(* IEC 61131-3 sources: Lasal-MCP/examples/SampleSource/2_PumpControlSolution/Stations/MachineControl/MachineControl/Class/SafetyBaseFSoE (part 3) *)

                b_NeedApplicationRestart := TRUE;
              end_if;
            end_if;
          end_if;
        end_if;

//*****************************************************************************
//**   UNSAFE BOOL INPUT VARIABLES                                           **
//*****************************************************************************

        // here we go for unsafe bool input vars

        // get number of unsafe input vars
        sd_retval := SDOReadCfgRequ ( p_SDORequestBuffer  := p_SDORequestBuffer
                                    , p_SDOResponseBuffer := p_SDOResponseBuffer
                                    , ud_Address          := ud_Address
                                    , us_Length           := 4
                                    );

        //no response
        if ( sd_retval <> 0 ) then
          LogError("@0217 (SafetyBaseFSoE::ReadSDOConfig) Config Read Error: Failed to read number of unsafe input vars.");
          return;
        end_if;

        ud_CntUnsafeInputs := p_SDOResponseBuffer^.ud_Data;

        ud_Address := p_SDORequestBuffer^.ud_Address + 4;

        // skip the names of unsafe inputs
        for i := 1 to ud_CntUnsafeInputs do

          // get length of Name
          sd_retval := SDOReadCfgRequ ( p_SDORequestBuffer  := p_SDORequestBuffer
                                      , p_SDOResponseBuffer := p_SDOResponseBuffer
                                      , ud_Address          := ud_Address
                                      , us_Length           := 4
                                      );
          //no response
          if ( sd_retval <> 0 ) then
            LogError("@0218 (SafetyBaseFSoE::ReadSDOConfig) Config Read Error: Reading length of unsafe input name failed.");
            return;
          end_if;

          // prepare address to get name
          ud_Address += 4;

//          ud_ActStrLen := ud_TmpStrLen := p_SDOResponseBuffer^.ud_Data;
          ud_TmpStrLen := p_SDOResponseBuffer^.ud_Data;
          ud_ActStrLen := ud_TmpStrLen;
          ud_TmpAddress := ud_Address;

          IF p_BlockedTransferMemory = NIL THEN
            sd_retval := -100;
            SetSafetyState(NewState:=_MemAllocFailed);
            RETURN;
          END_IF;

          IF ud_BlockedTransferMemorySize < (ud_TmpStrLen + 1) THEN
            p_BlockedTransferMemory := ToStdLib.ReAlloc(mptr:=p_BlockedTransferMemory, newsize:=GetNewMemSize(ud_TmpStrLen + 1));
            IF p_BlockedTransferMemory = NIL THEN
              ud_BlockedTransferMemorySize := 0;
              sd_retval := -100;
              SetSafetyState(NewState:=_MemAllocFailed);
              RETURN;
            ELSE
              ud_BlockedTransferMemorySize := GetNewMemSize(ud_TmpStrLen + 1);
            END_IF;
          END_IF;

          ToStdLib.MemSet(dest:=p_BlockedTransferMemory, value:=0, size:=ud_BlockedTransferMemorySize);

          p_TmpBlockedData := p_BlockedTransferMemory;

          us_BlockedTransferLength := BlockedTransferLength(ud_Datalength:=ud_TmpStrLen, us_MaxBlocklength:=60);

          while us_BlockedTransferLength do

            // get name
            sd_retval := SDOReadCfgRequ ( p_SDORequestBuffer  := p_SDORequestBuffer
                                        , p_SDOResponseBuffer := p_SDOResponseBuffer
                                        , ud_Address          := ud_TmpAddress
                                        , us_Length           := us_BlockedTransferLength
                                        , b_UseCache          := us_BlockedTransferLength < us_DataLength_Max
                                        );
            //no response
            if ( sd_retval <> 0 ) then
              LogError("@0219 (SafetyBaseFSoE::ReadSDOConfig) Config Read Error: Reading unsafe input name failed.");
              return;
            end_if;

            ToStdLib.MemCpy(dest:=p_TmpBlockedData,
                             source:=#p_SDOResponseBuffer^.ud_Data,
                             size:=us_BlockedTransferLength);

            p_TmpBlockedData += us_BlockedTransferLength;
            ud_TmpAddress += us_BlockedTransferLength;
            ud_TmpStrLen -= us_BlockedTransferLength;

            us_BlockedTransferLength := BlockedTransferLength(ud_Datalength:=ud_TmpStrLen, us_MaxBlocklength:=60);

          end_while;

          sd_retval := AddUnsafeRoutElement(pRoutTable:=#p_UnsafeInputsTable,
                                            pRoutElementsNo:=#ui_CntUnsafeInputs,
                                            ud_Address:=ud_ActAddress,
                                            ui_NameLen:=ud_ActStrLen$UINT,
                                            pNameNewElement:=p_BlockedTransferMemory$^CHAR);

          // if unsafe component not found (sd_retval <> 0), it's not problem for whole safe application

          // get offset in application memory
          ud_ActAddress += 4;

          // prepare address for next unsafe input
          ud_Address += ud_ActStrLen;

        end_for;

        // only available at new modules
        if b_CfgTypeV2 then

//*****************************************************************************
//**   UNSAFE BDINT INPUT VARIABLES                                          **
//*****************************************************************************

          // here we go for unsafe BDINT input vars

          // get number of unsafe input vars
          sd_retval := SDOReadCfgRequ ( p_SDORequestBuffer  := p_SDORequestBuffer
                                      , p_SDOResponseBuffer := p_SDOResponseBuffer
                                      , ud_Address          := ud_Address
                                      , us_Length           := 4
                                      );

          //no response
          if ( sd_retval <> 0 ) then
            LogError("@021A (SafetyBaseFSoE::ReadSDOConfig) Config Read Error: Failed to read number of unsafe BDINT input vars.");
            return;
          end_if;

          ud_CntUnsafeInputs := p_SDOResponseBuffer^.ud_Data;

          ud_Address := p_SDORequestBuffer^.ud_Address + 4;

          if ud_CntUnsafeInputs then

            //SDO request for this command has 5 bytes additional data
            pBitMasks$^void := ToStdLib.Malloc(size := ud_CntUnsafeInputs * sizeof(BDINT));

            if ( pBitMasks = NIL ) then
              sd_retval                         := -100;
              SetSafetyState(NewState:=_MemAllocFailed);
              LogError("@021B (SafetyBaseFSoE::ReadSDOConfig) Config Read Error: Failed to allocate memory for the BDINT variable bitmasks.");
              return;
            end_if;

            // get the bitmasks for the BDINT variables
            for i := 1 to ud_CntUnsafeInputs do

              // get bitmask
              sd_retval := SDOReadCfgRequ ( p_SDORequestBuffer  := p_SDORequestBuffer
                                          , p_SDOResponseBuffer := p_SDOResponseBuffer
                                          , ud_Address          := ud_Address
                                          , us_Length           := 4
                                          );
              //no response
              if ( sd_retval <> 0 ) then
                LogError("021C (SafetyBaseFSoE::ReadSDOConfig) Config Read Error: Reading bit mask of unsafe BDINT input failed.");
                return;
              end_if;

              // prepare address for the next one
              ud_Address += 4;

              // save the bitmask for adding the rout element
              (pBitMasks + (i-1) * sizeof(BDINT))^ := p_SDOResponseBuffer^.ud_Data;
            end_for;

            // get the names of unsafe inputs
            for i := 1 to ud_CntUnsafeInputs do

              // get length of Name
              sd_retval := SDOReadCfgRequ ( p_SDORequestBuffer  := p_SDORequestBuffer
                                          , p_SDOResponseBuffer := p_SDOResponseBuffer
                                          , ud_Address          := ud_Address
                                          , us_Length           := 4
                                          );
              //no response
              if ( sd_retval <> 0 ) then
                LogError("@021D (SafetyBaseFSoE::ReadSDOConfig) Config Read Error: Reading length of unsafe BDINT input name failed.");
                return;
              end_if;

              // prepare address to get name
              ud_Address += 4;

//              ud_ActStrLen := ud_TmpStrLen := p_SDOResponseBuffer^.ud_Data;
              ud_TmpStrLen := p_SDOResponseBuffer^.ud_Data;
              ud_ActStrLen := ud_TmpStrLen;
              ud_TmpAddress := ud_Address;

              IF p_BlockedTransferMemory = NIL THEN
                sd_retval := -100;
                SetSafetyState(NewState:=_MemAllocFailed);
                RETURN;
              END_IF;

              IF ud_BlockedTransferMemorySize < (ud_TmpStrLen + 1) THEN
                p_BlockedTransferMemory := ToStdLib.ReAlloc(mptr:=p_BlockedTransferMemory, newsize:=GetNewMemSize(ud_TmpStrLen + 1));
                IF p_BlockedTransferMemory = NIL THEN
                  ud_BlockedTransferMemorySize := 0;
                  sd_retval := -100;
                  SetSafetyState(NewState:=_MemAllocFailed);
                  RETURN;
                ELSE
                  ud_BlockedTransferMemorySize := GetNewMemSize(ud_TmpStrLen + 1);
                END_IF;
              END_IF;

              ToStdLib.MemSet(dest:=p_BlockedTransferMemory, value:=0, size:=ud_BlockedTransferMemorySize);

              p_TmpBlockedData := p_BlockedTransferMemory;

              us_BlockedTransferLength := BlockedTransferLength(ud_Datalength:=ud_TmpStrLen, us_MaxBlocklength:=60);

              while us_BlockedTransferLength do

                // get name
                sd_retval := SDOReadCfgRequ ( p_SDORequestBuffer  := p_SDORequestBuffer
                                            , p_SDOResponseBuffer := p_SDOResponseBuffer
                                            , ud_Address          := ud_TmpAddress
                                            , us_Length           := us_BlockedTransferLength
                                            , b_UseCache          := us_BlockedTransferLength < us_DataLength_Max
                                            );
                //no response
                if ( sd_retval <> 0 ) then
                  LogError("@021E (SafetyBaseFSoE::ReadSDOConfig) Config Read Error: Reading unsafe BDINT input name failed.");
                  return;
                end_if;

                ToStdLib.MemCpy(dest:=p_TmpBlockedData,
                                 source:=#p_SDOResponseBuffer^.ud_Data,
                                 size:=us_BlockedTransferLength);

                p_TmpBlockedData += us_BlockedTransferLength;
                ud_TmpAddress += us_BlockedTransferLength;
                ud_TmpStrLen -= us_BlockedTransferLength;

                us_BlockedTransferLength := BlockedTransferLength(ud_Datalength:=ud_TmpStrLen, us_MaxBlocklength:=60);

              end_while;

              ActBitMask := (pBitMasks + (i-1) * sizeof(BDINT))^;

              sd_retval := AddUnsafeRoutElement(pRoutTable:=#p_UnsafeInputsTable,
                                                pRoutElementsNo:=#ui_CntUnsafeInputs,
                                                ud_Address:=ud_UnsafeBDINT_Offset,
                                                ui_NameLen:=ud_ActStrLen$UINT,
                                                pNameNewElement:=p_BlockedTransferMemory$^CHAR,
                                                ActBitMask);

              // if unsafe component not found (sd_retval <> 0), it's not problem for whole safe application

              // get offset in application memory
              ud_ActAddress += CountBits(ActBitMask) * sizeof(DINT);
              ud_UnsafeBDINT_Offset += sizeof(DINT);

              // prepare address for next unsafe output or for number of constants
              ud_Address += ud_ActStrLen;

            end_for;

            // free the bitmasks
            ToStdLib.Free(mptr:=pBitMasks);
          end_if;

//*****************************************************************************
//**   CONSTANTS                                                             **
//*****************************************************************************

          // constants

          //send request and receive data
          sd_retval := SDOReadCfgRequ ( p_SDORequestBuffer  := p_SDORequestBuffer
                                      , p_SDOResponseBuffer := p_SDOResponseBuffer
                                      , ud_Address          := ud_Address
                                      , us_Length           := 4
                                      );

          //no response
          if ( sd_retval <> 0 ) then
            LogError("@021F (SafetyBaseFSoE::ReadSDOConfig) Config Read Error: Reading number of constants failed.");
            return;
          end_if;

          // skip number of constants
          ud_Address += 4;

          // skip constants
          ud_Address += p_SDOResponseBuffer^.ud_Data * 4;

          if b_CfgTypeV3 then

//*****************************************************************************
//**   SAFE DINT CONSTANTS                                                   **
//*****************************************************************************

            // constants

            //send request and receive data
            sd_retval := SDOReadCfgRequ ( p_SDORequestBuffer  := p_SDORequestBuffer
                                        , p_SDOResponseBuffer := p_SDOResponseBuffer
                                        , ud_Address          := ud_Address
                                        , us_Length           := 4
                                        );

            //no response
            if ( sd_retval <> 0 ) then
              LogError("@0220 (SafetyBaseFSoE::ReadSDOConfig) Config Read Error: Reading number of safe DINT constants failed.");
              return;
            end_if;

            // skip number of safe dint constants
            ud_Address += 4;

            // skip constants (4 byte per safe DINT constant)
            ud_Address += p_SDOResponseBuffer^.ud_Data * 4;

          end_if;

//*****************************************************************************
//**   LOCAL OUTPUTS                                                         **
//*****************************************************************************

          // local outputs
          //send request and receive data
          sd_retval := SDOReadCfgRequ ( p_SDORequestBuffer  := p_SDORequestBuffer
                                      , p_SDOResponseBuffer := p_SDOResponseBuffer
                                      , ud_Address          := ud_Address
                                      , us_Length           := 4
                                      );

          //no response
          if ( sd_retval <> 0 ) then
            LogError("@0221 (SafetyBaseFSoE::ReadSDOConfig) Config Read Error: Reading number of local outputs failed.");
            return;
          end_if;

          // skip number of local outputs
          ud_Address += 4;

          // skip local outputs
          //++pr
          // only available at new modules
          if b_CfgTypeV2 then
            ud_Address += p_SDOResponseBuffer^.ud_Data * 8; // Used-Flag, Modulkennung(SDIAS)
          else
            ud_Address += p_SDOResponseBuffer^.ud_Data * 4; // Used-Flag
          end_if;

          if b_CfgTypeV3 then

//*****************************************************************************
//**   LOCAL DINT OUTPUTS                                                    **
//*****************************************************************************

            // local outputs
            //send request and receive data
            sd_retval := SDOReadCfgRequ ( p_SDORequestBuffer  := p_SDORequestBuffer
                                        , p_SDOResponseBuffer := p_SDOResponseBuffer
                                        , ud_Address          := ud_Address
                                        , us_Length           := 4
                                        );

            //no response
            if ( sd_retval <> 0 ) then
              LogError("@0222 (SafetyBaseFSoE::ReadSDOConfig) Config Read Error: Reading number of local outputs failed.");
              return;
            end_if;

            // skip number of local outputs
            ud_Address += 4;

            // skip local outputs
            //++pr
            // only available at new modules
            if b_CfgTypeV2 then
              ud_Address += p_SDOResponseBuffer^.ud_Data * 8; // Used-Flag, Modulkennung(SDIAS)
            else
              ud_Address += p_SDOResponseBuffer^.ud_Data * 4; // Used-Flag
            end_if;

          end_if;

//*****************************************************************************
//**   SAFE BOOL INTERFACE OUTPUT VARIABLES                                  **
//*****************************************************************************

          // safe bool interface output vars
          //send request and receive data
          sd_retval := SDOReadCfgRequ ( p_SDORequestBuffer  := p_SDORequestBuffer
                                      , p_SDOResponseBuffer := p_SDOResponseBuffer
                                      , ud_Address          := ud_Address
                                      , us_Length           := 4
                                      );

          //no response
          if ( sd_retval <> 0 ) then
            LogError("@0223 (SafetyBaseFSoE::ReadSDOConfig) Config Read Error: Reading number of safe BOOL interface output variables failed.");
            return;
          end_if;

          // skip safe BOOL interface output variables
          ud_Address += 4;

          // count the interface output variables
          BoolOuts := p_SDOResponseBuffer^.ud_Data;

          if b_IsFSoE then
            ud_TmpCnt := p_SDOResponseBuffer^.ud_Data;

            if ud_TmpCnt then
              for i := 1 to ud_TmpCnt do
                //send request and receive data
                sd_retval := SDOReadCfgRequ ( p_SDORequestBuffer  := p_SDORequestBuffer
                                            , p_SDOResponseBuffer := p_SDOResponseBuffer
                                            , ud_Address          := ud_Address
                                            , us_Length           := 4
                                            );

                //no response
                if ( sd_retval <> 0 ) then
                  LogError("@027A (SafetyBaseFSoE::ReadSDOConfig) Config Read Error: Reading number of FSoE connections for BOOL interface outputs failed.");
                  return;
                end_if;

                // skip number of entries and the entries
                ud_Address += 4 + 4 * p_SDOResponseBuffer^.ud_Data;
              end_for;
            end_if;
          end_if;

//*****************************************************************************
//**   SAFE DINT INTERFACE OUTPUT VARIABLES                                  **
//*****************************************************************************

          // safe dint interface output vars
          //send request and receive data
          sd_retval := SDOReadCfgRequ ( p_SDORequestBuffer  := p_SDORequestBuffer
                                      , p_SDOResponseBuffer := p_SDOResponseBuffer
                                      , ud_Address          := ud_Address
                                      , us_Length           := 4
                                      );

          //no response
          if ( sd_retval <> 0 ) then
            LogError("@0224 (SafetyBaseFSoE::ReadSDOConfig) Config Read Error: Reading number of safe DINT interface output variables failed.");
            return;
          end_if;

          // skip number of safe dint interface output vars
          ud_Address += 4;

          // count the interface output variables
          DintOuts := p_SDOResponseBuffer^.ud_Data;

          if b_IsFSoE then
            ud_TmpCnt := p_SDOResponseBuffer^.ud_Data;

            if ud_TmpCnt then
              for i := 1 to ud_TmpCnt do
                //send request and receive data
                sd_retval := SDOReadCfgRequ ( p_SDORequestBuffer  := p_SDORequestBuffer
                                            , p_SDOResponseBuffer := p_SDOResponseBuffer
                                            , ud_Address          := ud_Address
                                            , us_Length           := 4
                                            );

                //no response
                if ( sd_retval <> 0 ) then
                  LogError("@027B (SafetyBaseFSoE::ReadSDOConfig) Config Read Error: Reading number of FSoE connections for DINT interface outputs failed.");
                  return;
                end_if;

                // skip number of entries and the entries
                ud_Address += 4 + 4 * p_SDOResponseBuffer^.ud_Data;
              end_for;
            end_if;
          end_if;

//*****************************************************************************
//**   FSBs = Functional Safety Blocks                                       **
//*****************************************************************************

          ud_skipLength := 0;

          // skip FSBs! structure: CRC, Length.... until the length is 0
          repeat

            // skip CRC and length of FSB
            ud_Address += 4 + ud_skipLength;

            //send request and receive data
            sd_retval := SDOReadCfgRequ ( p_SDORequestBuffer  := p_SDORequestBuffer
                                        , p_SDOResponseBuffer := p_SDOResponseBuffer
                                        , ud_Address          := ud_Address
                                        , us_Length           := 4
                                        );

            //no response
            if ( sd_retval <> 0 ) then
              LogError("@0225 (SafetyBaseFSoE::ReadSDOConfig) Config Read Error: Reading length of FSB failed.");
              return;
            end_if;

            ud_skipLength := p_SDOResponseBuffer^.ud_Data;

          until ud_skipLength = 0 end_repeat;

          // skip length of block with 0 length
          ud_Address += 4;

          if b_CfgTypeV3 then

//*****************************************************************************
//**   DYNAMIC PARAMETERS (e.g. for SSI Module)                              **
//*****************************************************************************

// Version of Parameters is saved in hd_DynParaVersion
// if it's 16#0001, then we read out the number of parameters which will follow

// structure:
// number of parameters
// for every parameter: place, id, length (including the 4 byte for the length itself), data

            //send request and receive data
            sd_retval := SDOReadCfgRequ ( p_SDORequestBuffer  := p_SDORequestBuffer
                                        , p_SDOResponseBuffer := p_SDOResponseBuffer
                                        , ud_Address          := ud_Address
                                        , us_Length           := 4
                                        );

            //no response
            if ( sd_retval <> 0 ) then
              LogError("@0226 (SafetyBaseFSoE::ReadSDOConfig) Config Read Error: Reading number of dynamic parameters failed.");
              return;
            end_if;

            ud_TmpCnt := p_SDOResponseBuffer^.ud_Data;

            // skip number of parameters
            ud_Address += 4;

            if ud_TmpCnt then
              for i := 1 to ud_TmpCnt do
                //send request and receive data
                sd_retval := SDOReadCfgRequ ( p_SDORequestBuffer  := p_SDORequestBuffer
                                            , p_SDOResponseBuffer := p_SDOResponseBuffer
                                            , ud_Address          := ud_Address
                                            , us_Length           := sizeof(t_DynamicParameterHeader)
                                            );

                //no response
                if ( sd_retval <> 0 ) then
                  LogError("@0227 (SafetyBaseFSoE::ReadSDOConfig) Config Read Error: Reading header of dynamic parameter failed.");
                  return;
                end_if;

                DynamicParameterHeader := p_SDOResponseBuffer^.ud_Data$t_DynamicParameterHeader;

                AddressServiceDataSize := 0;

                // skip size of header
                ud_Address += sizeof(t_DynamicParameterHeader);

                // data for pdo length info:
                // this data is also mirrored to SBF_SDO_ADDRESS_SPECIAL_INFO

//                  Marked with Place = 1000
//
//                  (4 Byte Length)
//                   4 Byte Version (starting at 0)
//                   1 Byte Length Rd PDO
//                   1 Byte Length Rd PDO IF
//                   1 Byte Length Wr PDO
//                   1 Byte Number of write PDOs (without additional it would be 1), msb = fast unsafe active

                if (DynamicParameterHeader.Place = SBF_CONFIG_PDO_INFO_PLACE) & (DynamicParameterHeader.Length >= (sizeof(UDINT) + sizeof(t_PDOSizeInfo))) then
                  //send request and receive data
                  sd_retval := SDOReadCfgRequ ( p_SDORequestBuffer  := p_SDORequestBuffer
                                              , p_SDOResponseBuffer := p_SDOResponseBuffer
                                              , ud_Address          := ud_Address
                                              , us_Length           := sizeof(t_PDOSizeInfo)
                                              );

                  //no response
                  if ( sd_retval <> 0 ) then
                    LogError("@0228 (SafetyBaseFSoE::ReadSDOConfig) Config Read Error: Reading dynamic parameter for pdo size failed.");
                    return;
                  end_if;

                  ud_Address += sizeof(t_PDOSizeInfo);

                  AddressServiceDataSize := (ud_ListLength_Address + ud_ListLength) - ud_Address;

                  PdoSizeInfo := p_SDOResponseBuffer^.ud_Data$t_PDOSizeInfo;

                  // if any sizes increased or we would need more DOs
                  if (PdoSizeInfo.PDORdLen > MyPDOReadSize)     |
                     (PdoSizeInfo.PDOWrLen > MyPDOWriteSize)    |
                     ((PdoSizeInfo.FastUnsafeAvailable <> 0) > ActivateFastUnsafeIOs) then

                    // error => can't go on like this
                    LogError("@0202 (SafetyBaseFSoE::ReadSDOConfig) Number or size of module accesses increased with new safety project!");
                    LogError("@0203 (SafetyBaseFSoE::ReadSDOConfig) => Can't continue, because the new data is not covered by the actual accesses! Restart Application!");

                    b_NeedApplicationRestart := TRUE;
                  end_if;

                  exit;
                end_if;

                // skip the parameter data (length of the length is also included)
                ud_Address += DynamicParameterHeader.Length - 4;
              end_for;

              if AddressServiceDataSize then
(*

  Data structure of address service data

  4 Byte Anzahl der MultiChannel
    Pro MultiChannel:
    4 Byte Anzahl der Verwendungen des Multichannel
    4 Byte Index des Gesamtergebnisses
    1 Byte Art der Verknüpfung (0 = UND)
    1 Byte Defaultbelegung des Werts
    2 Byte Reserved (für 4 Byte Alignment)
      Pro Verwendung (siehe erster Eintrag in den MultiChannelDaten):
      4 Byte FSoE Daten
  4 Byte Kommunikations-ID (Default 0)
  4 Byte Anzahl der Adressbereiche
    Pro Adressbereich:
    4 Byte Startadresse
    4 Byte Länge Adressbereich
  4 Byte Anzahl der Connection-ID-Bereiche
    Pro Bereich:
    4 Byte Startadresse
    4 Byte Länge Bereich

*)
                // get the number of multichannels
                sd_retval := SDOReadCfgRequ ( p_SDORequestBuffer  := p_SDORequestBuffer
                                            , p_SDOResponseBuffer := p_SDOResponseBuffer
                                            , ud_Address          := ud_Address
                                            , us_Length           := 4
                                            );

                //no response
                if ( sd_retval <> 0 ) then
                  LogError("@027C (SafetyBaseFSoE::ReadSDOConfig) Config Read Error: Reading address service data failed.");
                  return;
                end_if;

                ud_TmpCnt := p_SDOResponseBuffer^.ud_Data;

                // skip number of multichannels
                ud_Address += 4;

                if ud_TmpCnt then
                  for i := 1 to ud_TmpCnt do
                    // get the number of usages
                    sd_retval := SDOReadCfgRequ ( p_SDORequestBuffer  := p_SDORequestBuffer
                                                , p_SDOResponseBuffer := p_SDOResponseBuffer
                                                , ud_Address          := ud_Address
                                                , us_Length           := 4
                                                );

                    //no response
                    if ( sd_retval <> 0 ) then
                      LogError("@027C (SafetyBaseFSoE::ReadSDOConfig) Config Read Error: Reading address service data failed.");
                      return;
                    end_if;

                    // skip the rest of this multichannel
                    ud_Address += 12 + (p_SDOResponseBuffer^.ud_Data * 4);
                  end_for;
                end_if;

                // skip the communication ID
                ud_Address += 4;

                // read the number of address areas
                sd_retval := SDOReadCfgRequ ( p_SDORequestBuffer  := p_SDORequestBuffer
                                            , p_SDOResponseBuffer := p_SDOResponseBuffer
                                            , ud_Address          := ud_Address
                                            , us_Length           := 4
                                            );

                //no response
                if ( sd_retval <> 0 ) then
                  LogError("@027C (SafetyBaseFSoE::ReadSDOConfig) Config Read Error: Reading address service data failed.");
                  return;
                end_if;

                // if there are any => the module got an address service
                if p_SDOResponseBuffer^.ud_Data then
                  TempModuleConfig.Info.IsAddressService := TRUE;
                end_if;
              end_if;
            end_if;
          end_if;

          // if there are interface variables
          if BoolOuts | DintOuts then
            // calculate the length of the interface frame
            TempPdoConfig.PdoLen := CalcPDOLength(BoolOuts, DintOuts);

            TempPdoConfig.Info := 0;
            TempPdoConfig.Info.IsInterfacePDO := TRUE;
            TempPdoConfig.Info.IsOptional := (ud_ActBlockType = SBF_BLKTYPE_CFG_MODULE_OPTIONAL);

            // if it's a broadcast => mark it
            if (TempPath[0]$UINT = 2) & (TempPath[0]$HDINT = SBF_INTERFACE_FRAME_BROADCAST) then
              TempPdoConfig.Info.IFBroadCast := TRUE;
            end_if;

            // this is the source of the interface frame
            TempPdoConfig.SourcePathLen := pListHeader^.p_us_Path^$UINT + 2;
            TempPdoConfig.pSourcePath   := pListHeader^.p_us_Path;

            // and the destination
            TempPdoConfig.DestPathLen   := TempPath[0]$UINT + 2;
            TempPdoConfig.pDestPath     := #TempPath[0];

            // add the interface PDO to the list
//            AddPdoToCfg(TempPdoConfig);

            TempModuleConfig.Info.IsInterfaceSource := TRUE;
            TempModuleConfig.Info.IsInterfaceDest   := FALSE;
            TempModuleConfig.InterfaceCRC := TempPdoConfig.InterfaceCRC;
          else
            TempModuleConfig.Info.IsInterfaceSource := FALSE;
            TempModuleConfig.Info.IsInterfaceDest   := FALSE;
            TempModuleConfig.InterfaceCRC := 0;
          end_if;
        else
          TempModuleConfig.Info.IsInterfaceSource := FALSE;
          TempModuleConfig.Info.IsInterfaceDest   := FALSE;
          TempModuleConfig.InterfaceCRC := 0;
        end_if;

        // if it's our own path, remember the safety number
        if (PathOfThisCPU[0]$UINT = (pListHeader^.p_us_Path$^UINT)^) & (ToStdLib.MemCmp(#PathOfThisCPU[0], pListHeader^.p_us_Path, PathOfThisCPU[0]$UINT + 2) = 0) then
          TempModuleConfig.SafetyNbr := SafetyNumber;
          //safe config of scp modul (own path)
          SafeActModuleConfig(TempModuleConfig);
        else
          TempModuleConfig.SafetyNbr := 0;
        end_if;

        // only when there is a manager
        if pSafetyManagerThis then
          AddModuleToCfg(TempModuleConfig);
        end_if;

//**********************************************************************************************************************************************************
      SBF_BLKTYPE_OLD_MODE_FLAG: // flag fore FW to use old config-mode
        // we need the old TimeSync config-type
        NewConfigType := ConfigState_Old;

//**********************************************************************************************************************************************************
      SBF_BLKTYPE_CFG_XML: // configuration for uploading the project to the safetydesigner (network placement information, names of bits,...)
        // no useful information here for us

//**********************************************************************************************************************************************************
    else
      // skip it = do nothing
//      TRACE("Found unhandled Blocktype in configuration.");
//**********************************************************************************************************************************************************
    end_case;

    ud_ListBaseAddress := ud_ListLength_Address + ud_ListLength;
  end_while;

  if ( ( sd_retval = 0 ) & ( SafetyState = _ModFromCfgNotFound ) ) then
    sd_retval := -1;
  end_if;

END_FUNCTION

FUNCTION VIRTUAL SafetyBaseFSoE::SDOReadCfgRequ
  VAR_INPUT
    p_SDORequestBuffer 	: ^SafetyBaseFSoE::SDORequReadConfig;
    p_SDOResponseBuffer 	: ^SafetyBaseFSoE::SDORespReadConfig;
    ud_Address 	: UDINT;
    us_Length 	: USINT;
    b_UseCache 	: BOOL;(* := TRUE *)
  END_VAR
  VAR_OUTPUT
    sd_retval 	: DINT;
  END_VAR

  // check if we have the data in the cache
  if b_UseCache & IsInCache(ud_Address, us_Length) then
    // use it from the cache

    // the address may be used from outside this function
    p_SDORequestBuffer^.ud_Address := ud_Address;

    _memcpy(ptr1:=#p_SDOResponseBuffer^.ud_Data, ptr2:=#Cache[0] + (ud_Address - CachedAddr), cntr:=us_Length);

    // everything is fine
    sd_retval := 0;
  else

    //sequence number
    p_SDORequestBuffer^.StdHeader.SeqNr := us_CntSequNr;

    //increase counter for sequence number
    if us_CntSequNr < 16#7F then
      us_CntSequNr += 1;
    else
      us_CntSequNr := 0;
    end_if;

    //address
    p_SDORequestBuffer^.ud_Address := ud_Address;

    if b_UseCache then
      // get max size
      p_SDORequestBuffer^.us_Length := SBF_SDO_MAX_LENGTH - (sizeof(SDORespReadConfig) - sizeof(SDORespReadConfig.ud_Data));
    else
      //length of expected data
      p_SDORequestBuffer^.us_Length := us_Length;
    end_if;

    //calculate CRC (starting with length of data until the end of command)
    p_SDORequestBuffer^.StdHeader.CRC := 0;

    //send request
    sd_retval := SAFETY_iSendRequest( uiMaster    := 0
                                    , pucNode     := p_ObjectPath
                                    , uiInLength  := sizeof(SDORequReadConfig)
                                    , pucInput    := p_SDORequestBuffer$^USINT
                                    , uiOutLength := sizeof(SDORespReadConfig) - sizeof(SDORespReadConfig.ud_Data) + p_SDORequestBuffer^.us_Length
                                    , pucOutput   := p_SDOResponseBuffer$^USINT
                                    );

    //no response
    if ( sd_retval <> 0 ) then
      LogError("@0229 (SafetyBaseFSoE::SDOReadCfgRequ) SAFETY_iSendRequest failed.");

      // we remember to retry in a few seconds
      b_ReadConfigFailed := TRUE;
      return;
    end_if;

    //check sequence number to exclude a possible wrong response
    if ( p_SDORequestBuffer^.StdHeader.SeqNr <> p_SDOResponseBuffer^.StdHeader.SeqNr ) then
      // we remember to retry in a few seconds
      b_ReadConfigFailed := TRUE;
      //log not routable SDOs
      LogValue("@022A (SafetyBaseFSoE::SDOReadCfgRequ) Invalid Sequence number in SDO Standard Response. Got 0x{0} instead of expected 0x{1}", to_udint(p_SDOResponseBuffer^.StdHeader.SeqNr), to_udint(p_SDORequestBuffer^.StdHeader.SeqNr));
      return;
    end_if;

    //check returncode of SDO
    if ( p_SDOResponseBuffer^.us_Returncode <> SBF_SDO_RETCODE_OK ) then
      //log not routable SDOs
      LogValue("@022B (SafetyBaseFSoE::SDOReadCfgRequ) Safety module 0x{0}: Retcode of SDO Standard Response was invalid. Retcode: 0x{1}", SafetyNumber$UDINT, to_udint(p_SDOResponseBuffer^.us_Returncode));

  //    // when reading fails because safety designer is writing at the same moment
  //    if p_SDOResponseBuffer^.us_Returncode = SDO_MICROCTRL_DIFFER then
        // we remember to retry in a few seconds
        b_ReadConfigFailed := TRUE;
  //    end_if;

      return;
    end_if;

    //check length of read data
    if ( p_SDOResponseBuffer^.us_Length = 0 ) then
      LogError("@022C (SafetyBaseFSoE::SDOReadCfgRequ) Response length is 0.");
      sd_retval := -104;
      return;
    elsif b_UseCache then
      // everything is fine => add the new data to the cache
      AddToCache(p_SDORequestBuffer, p_SDOResponseBuffer);
    end_if;
  end_if;

END_FUNCTION

FUNCTION VIRTUAL SafetyBaseFSoE::GetRoutingData
  VAR_OUTPUT
    sd_retval 	: DINT;
  END_VAR
  VAR
    SDORequestBuffer        : SDORequReadConfig;
    SDOResponseBuffer       : ARRAY [0..SBF_SDO_MAX_LENGTH-1] OF USINT;
    p_SDORequestBuffer 	    : ^SDORequReadConfig;
    p_SDOResponseBuffer 	  : ^SDORespReadConfig;
    Module                  : PathInfoType;
    ListHeader              : PathInfoType;
    NotAvailableStr         : ARRAY [0..99] OF CHAR;
    ModulePath              : ARRAY [0..127] OF USINT;
    ModulePathComp          : ARRAY [0..127] OF USINT;
    ListPath                : ARRAY [0..127] OF USINT;
    ListPathComp            : ARRAY [0..127] OF USINT;
    Time1, Time2            : UDINT;
  END_VAR

  // get module specific configuration information
  GetConfiguration();

  InitPathInfo(#Module);
  InitPathInfo(#ListHeader);

  //SDO request for this command has 5 bytes additional to the header
  p_SDORequestBuffer := #SDORequestBuffer;

  //SDO response for this command can have maximum additional data
  p_SDOResponseBuffer := (#SDOResponseBuffer)$^SDORespReadConfig;

  //path of input-safety-module
  Module.p_us_Path$^void := #ModulePath;

  //compressed path of input-safety-module
  Module.p_us_PathComp$^void := #ModulePathComp;

  //path in list header
  ListHeader.p_us_Path$^void := #ListPath;

  //path in list header
  ListHeader.p_us_PathComp$^void := #ListPathComp;

  b_ReadConfigFailed := FALSE;

  b_NeedApplicationRestart := FALSE;

  // if there is a revision in the configuration this variable changes to TRUE
  b_GotNewRevision := FALSE;

Time1 := OS_READMICROSEC();
  //read config data via SDOs and add safety modules to routing lists
  sd_retval := ReadSDOConfig( p_SDORequestBuffer      := p_SDORequestBuffer
                            , p_SDOResponseBuffer     := p_SDOResponseBuffer
                            , pModule                 := #Module
                            , pListHeader             := #ListHeader
                            );
Time2 := OS_READMICROSEC();
ud_ConfigReadTime := Time2 - Time1;

  // set error to restart application afterwards to have a complete configuration (needed for routing to share the slave configurations with only 1 restart of the application)
  if b_NeedApplicationRestart then
    SetSafetyState(NewState:=_DOsIncreasedRestartApp);
    sd_retval := -1;
  end_if;

  // if there is no revision in the configuration => clear it
  if (b_GotNewRevision = FALSE) then

    // free memory, if available
    if pPrjNameStr & pPrjRevStr then
      ToStdLib.Free(pPrjNameStr);
    end_if;

    // use local memory to show "not available"
    _strcpy(dest:=#NotAvailableStr[0], src:="<not available>");
    PrjNameMemLen := _strlen(src:=#NotAvailableStr[0]);
    PrjNameStrLen := PrjRevStrLen := PrjNameMemLen - 1;
    pPrjNameStr := pPrjRevStr := #NotAvailableStr[0];

    // write the strings to the string objects
    ShowProjectRevision();

    // there is no memory, so reset the pointer and length informations
    pPrjNameStr := NIL;
    pPrjRevStr := NIL;

    PrjNameMemLen := 0;
    PrjNameStrLen := 0;
    PrjRevStrLen := 0;
  end_if;

  // if reading failed, because designer is writing at the same time => we try again in a few seconds
  if b_ReadConfigFailed then

    // next time we check for the configured state of the cpu
    b_CheckConfigured := TRUE;

    // check again in background
    SetSafetyState(NewState:=_ReinitConfig);

    // and wait at least 3 secs
    ud_LastCheckConfig := ops.tAbsolute;

  // error in configuration -> no work
  elsif ( sd_retval <> 0 ) & (SafetyState <> _ReinitConfig) then
    if SafetyState = _WaitForSynchronicity then
      SetSafetyState(NewState:=_UnknownCfgError);
    end_if;

    LogError("@022D (SafetyBaseFSoE::GetRoutingData) Reading Safety Configuration failed!");
  else
    // read config succeeded, check update cycle of unsafe variables
    CheckUnsafeUpdateCycle();

    // check for interface frame destination modules and mark them
    GetDestinationCRCs();

    // if there is a safety manager create a configuration message and send it to the safety manager
    if pSafetyManagerThis then
      CreateAndSendCfg();
    end_if;

    // last thing to do is to start realtime and cyclic work (they do nothing in _ReinitConfig state
    if ud_UnsafeVarsNotFound then
      SetSafetyState(NewState:=_UnsafeVarNotFound);
      ud_UnsafeVarsNotFound := 0;
    else
      if us_SetBusReadyState = SetBusReadyFinished then
        // we're already synchron from a former configuration phase
        SetSafetyState(NewState:=_SafetyClassOK);
      else
        SetSafetyState(NewState:=_WaitForSynchronicity);
      end_if;
    end_if;
  end_if;

  // free temporary configuration lists if there were any
  FreeCfgLists();

END_FUNCTION

FUNCTION VIRTUAL SafetyBaseFSoE::ReadModulePath
  VAR_INPUT
    p_SDORequestBuffer 	: ^SafetyBaseFSoE::SDORequReadConfig;
    p_SDOResponseBuffer 	: ^SafetyBaseFSoE::SDORespReadConfig;
    p_ud_Address 	: ^UDINT;
    pModule 	: ^SafetyBaseFSoE::PathInfoType;
    p_ud_ModulePathLen_Max 	: ^UDINT;
    p_ud_ModulePathCompLen_Max 	: ^UDINT;
    us_SDOMaxDataSize 	: USINT;
  END_VAR
  VAR_OUTPUT
    sd_retval 	: DINT;
  END_VAR
  VAR
    ud_ModulePathLen_Act    : UDINT;
    p_ud_ModulePath_Act     : ^UDINT;
  END_VAR

  //read length of module path

  //send request and receive data
  sd_retval := SDOReadCfgRequ ( p_SDORequestBuffer  := p_SDORequestBuffer
                              , p_SDOResponseBuffer := p_SDOResponseBuffer
                              , ud_Address          := p_ud_Address^
                              , us_Length           := 4
                              );

  //no response
  if ( sd_retval <> 0 ) then
    LogError("@022E (SafetyBaseFSoE::ReadModulePath) Failed to read length of module path.");
    return;
  end_if;

  //length of module path
  ud_ModulePathLen_Act := p_SDOResponseBuffer^.ud_Data;

  //length is zero, check compressed path
  if ( ud_ModulePathLen_Act > 0 ) then

    // if it's too small => error
    if ( ud_ModulePathLen_Act > p_ud_ModulePathLen_Max^ ) then
      sd_retval                         := -100;
      SetSafetyState(NewState:=_MemAllocFailed);
      return;
    end_if;

    //read path

    //address of first byte of path
    p_ud_Address^ += 4;

    //set pointer to first byte of target buffer
    p_ud_ModulePath_Act := ( pModule^.p_us_Path )$^UDINT;

    //read path block by block, if path is longer than max. length
    while ( ud_ModulePathLen_Act > us_SDOMaxDataSize ) do

      //send request and receive data
      sd_retval := SDOReadCfgRequ ( p_SDORequestBuffer  := p_SDORequestBuffer
                                  , p_SDOResponseBuffer := p_SDOResponseBuffer
                                  , ud_Address          := p_ud_Address^
                                  , us_Length           := us_SDOMaxDataSize
                                  , b_UseCache          := FALSE
                                  );

      //no response
      if ( sd_retval <> 0 ) then
        LogError("@022F (SafetyBaseFSoE::ReadModulePath) Failed to read block of module path.");
        return;
      end_if;

      //copy part of path
      ToStdLib.MemCpy(dest := p_ud_ModulePath_Act , source := #p_SDOResponseBuffer^.ud_Data, size := us_SDOMaxDataSize);

      //rest of path to be read
      ud_ModulePathLen_Act -= us_SDOMaxDataSize;

      //address of next block
      p_ud_Address^ += us_SDOMaxDataSize;

      //set pointer to next free byte of target buffer
      p_ud_ModulePath_Act += us_SDOMaxDataSize;

    end_while;

    // if there is something left
    if ud_ModulePathLen_Act then
      //read last bytes of path

      //send request and receive data
      sd_retval := SDOReadCfgRequ ( p_SDORequestBuffer  := p_SDORequestBuffer
                                  , p_SDOResponseBuffer := p_SDOResponseBuffer
                                  , ud_Address          := p_ud_Address^
                                  , us_Length           := ud_ModulePathLen_Act$USINT
                                  , b_UseCache          := ud_ModulePathLen_Act$USINT < us_SDOMaxDataSize
                                  );

      //no response
      if ( sd_retval <> 0 ) then
        LogError("@0230 (SafetyBaseFSoE::ReadModulePath) Failed to read last bytes of module path.");
        return;
      end_if;

      ToStdLib.MemCpy(dest := p_ud_ModulePath_Act, source := #p_SDOResponseBuffer^.ud_Data, size := ud_ModulePathLen_Act);
    end_if;

    //address of next byte after path
    //address of last block + length of last read block
    p_ud_Address^ += ud_ModulePathLen_Act;
  else
    pModule^.p_us_Path := NIL;

    //address of compressed path
    p_ud_Address^ += 4;
  end_if;

// ============================================================================================================================

  // compressed module path starts here

  // read length of module path

  // send request and receive data
  sd_retval := SDOReadCfgRequ ( p_SDORequestBuffer  := p_SDORequestBuffer
                              , p_SDOResponseBuffer := p_SDOResponseBuffer
                              , ud_Address          := p_ud_Address^
                              , us_Length           := 4
                              );

  //no response
  if ( sd_retval <> 0 ) then
    LogError("@0231 (SafetyBaseFSoE::ReadModulePath) Failed to read length of compressed module path.");
    return;
  end_if;

  //length of module path
  ud_ModulePathLen_Act := p_SDOResponseBuffer^.ud_Data;

  pModule^.ui_PathCompLen := to_uint(ud_ModulePathLen_Act);

  //if length is zero, leave method
  if ( ud_ModulePathLen_Act = 0 ) then
    if pModule^.p_us_PathComp <> NIL then
      pModule^.p_us_PathComp := NIL;
    end_if;

    // address of CRC
    p_ud_Address^ += 4;

    return;
  end_if;

  //if it's too small => error
  if ( ud_ModulePathLen_Act > p_ud_ModulePathCompLen_Max^ ) then
    sd_retval                         := -100;
    SetSafetyState(NewState:=_MemAllocFailed);
    return;
  end_if;

  //read path

  //address of first byte of path
  p_ud_Address^ += 4;

  //set pointer to first byte of target buffer
  p_ud_ModulePath_Act := pModule^.p_us_PathComp$^UDINT;

  //read path block by block, if path is longer than max. length
  while ( ud_ModulePathLen_Act > us_SDOMaxDataSize ) do

    //send request and receive data
    sd_retval := SDOReadCfgRequ ( p_SDORequestBuffer  := p_SDORequestBuffer
                                , p_SDOResponseBuffer := p_SDOResponseBuffer
                                , ud_Address          := p_ud_Address^
                                , us_Length           := us_SDOMaxDataSize
                                , b_UseCache          := FALSE
                                );

    //no response
    if ( sd_retval <> 0 ) then
      LogError("@0232 (SafetyBaseFSoE::ReadModulePath) Failed to read block of compressed module path.");
      return;
    end_if;

    //copy part of path
    ToStdLib.MemCpy(dest := p_ud_ModulePath_Act , source := #p_SDOResponseBuffer^.ud_Data, size := us_SDOMaxDataSize);

    //rest of path to be read
    ud_ModulePathLen_Act -= us_SDOMaxDataSize;

    //address of next block
    p_ud_Address^ += us_SDOMaxDataSize;

    //set pointer to next free byte of target buffer
    p_ud_ModulePath_Act += us_SDOMaxDataSize;

  end_while;

  // if there is something left
  if ud_ModulePathLen_Act then

    //read last bytes of path

    //send request and receive data
    sd_retval := SDOReadCfgRequ ( p_SDORequestBuffer  := p_SDORequestBuffer
                                , p_SDOResponseBuffer := p_SDOResponseBuffer
                                , ud_Address          := p_ud_Address^
                                , us_Length           := ud_ModulePathLen_Act$USINT
                                , b_UseCache          := ud_ModulePathLen_Act$USINT < us_SDOMaxDataSize
                                );

    //no response
    if ( sd_retval <> 0 ) then
      LogError("@0233 (SafetyBaseFSoE::ReadModulePath) Failed to read last bytes of compressed module path.");
      return;
    end_if;

    ToStdLib.MemCpy(dest := p_ud_ModulePath_Act, source := #p_SDOResponseBuffer^.ud_Data, size := ud_ModulePathLen_Act);
  end_if;

  //address of next byte after path
  //address of last block + length of last read block
  p_ud_Address^ += ud_ModulePathLen_Act;

END_FUNCTION

FUNCTION VIRTUAL SafetyBaseFSoE::AddModuleToRoutingTabs
  VAR_INPUT
    pModule 	: ^SafetyBaseFSoE::PathInfoType;
    pListHeader 	: ^SafetyBaseFSoE::PathInfoType;
    b_IsOptional 	: BOOL;
  END_VAR
  VAR_OUTPUT
    sd_retval 	: DINT;
  END_VAR
  VAR
    p_TargetObject            : pVirtualBase;
    p_SafetyBase              : pVirtualBase;
    ud_IO_SafeNumber          : HDINT;
    ud_PDO_Buffer             : UDINT;
    MyPara 	                  : CmdStruct;
    MyResult	                : results;
  END_VAR

//#pragma message("RamAnd 29.10.2014 10:26 \ hier kann vermutlich config in/out/cpu entfallen. einfach nur die entsprechenden module merken")

  //get this-pointer of object in network that is located with transfered path
  MyPara.uiCmd := _BUS_IF_GET_OBJECT_THIS_PTR;
  MyPara.aPara[0] := pModule^.p_us_Path$DINT;
  sd_retval$iprStates := ToBusInterface.NewInst(#MyPara, #MyResult);
  p_TargetObject := MyResult.aData[0]$pVirtualBase;

  //this-pointer found
  if ( p_TargetObject ) then

    //add output module

    //If found this-pointer equals the own this-pointer, then the module has to be added to output-list.
    //This module (CPU) provides the safety input values for the output module (path in list-header).
    if ( p_TargetObject = this ) then

      //the output module is addressed by the ListHeaderPath
      //get this-pointer of object in network that is located with transfered path
      MyPara.uiCmd := _BUS_IF_GET_OBJECT_THIS_PTR;
      MyPara.aPara[0] := pListHeader^.p_us_Path$DINT;
      sd_retval$iprStates := ToBusInterface.NewInst(#MyPara, #MyResult);
      p_TargetObject := MyResult.aData[0]$pVirtualBase;

      //this-pointer found
      if ( p_TargetObject ) then

        MyPara.uiCmd := CMD_SM_GET_MODULE_TYPE;
        sd_retval$iprStates := p_TargetObject^.NewInst(#MyPara, #MyResult);

        //check if it's a safety module with FSoE
        if ( MyResult.aData[0]$UDINT = SM_TYPE_SAFETY_MODULE_FSOE ) then

          //object is based on SafetyBaseFSoE
          p_SafetyBase := ( p_TargetObject )$pVirtualBase;

          //get pointer on PDO output buffer
          ud_PDO_Buffer := GetPointer2PDOBuffer();

          //configure safety output module and receive safety number
          //inform the output module about safety number and object path of the safe CPU

          //get safety number
          MyPara.uiCmd := CMD_SM_CONFIG_SAFETY_CPU;

          sd_retval$iprStates := p_SafetyBase^.NewInst(#MyPara, #MyResult);

          ud_IO_SafeNumber := MyResult.aData[0]$UDINT;
//
//          MyPara.uiCmd := CMD_SM_CONFIG_SAFETY_OUTPUT;
//          MyPara.aPara[0] := SafetyNumber$DINT;
//          MyPara.aPara[1] := this$DINT;
//          MyPara.aPara[2] := (GetPointer2PDOBuffer())$DINT;
//          MyPara.aPara[3] := pModule$DINT;
//          MyPara.aPara[6] := b_IsOptional;
//          MyPara.aPara[7] := 0; // Pass DO Handle           p_HandlePDORead$DINT;
//          MyPara.aPara[8] := 0; // Offset within the DO     0$DINT;
//
//          sd_retval$iprStates := p_SafetyBase^.NewInst(#MyPara, #MyResult);
//
//          ud_IO_SafeNumber := MyResult.aData[0]$UDINT;

//          ud_IO_SafeNumber := p_SafetyBase^.ConfigSafetyOutput  ( ud_SafeNrCPU    := SafetyNumber
//                                                                , ud_thisp        := this$UDINT
//                                                                , ud_p_PDOBuffer  := GetPointer2PDOBuffer()
//                                                                , pObject         := pModule
//                                                                , pMoveActive     := pMoveCommandOutputActive
//                                                                , ud_MoveSourceAddr := ud_LocalMoveSourceAddr
//                                                                , b_IsOptional := b_IsOptional
//                                                                );

          //output module successfully configured
          if ( ud_IO_SafeNumber <> 0 ) then

            //add module to routing table
            sd_retval := AddRoutingElement( ud_SafeNumber       := ud_IO_SafeNumber
                                          , ud_thisp            := p_SafetyBase$UDINT
                                          , pObject             := pListHeader
                                          );
          else
            sd_retval := 0; // could be an optional module
          end_if;
        else
          LogError("@027D (SafetyBaseFSoE::AddModuleToRoutingTabs) Config Read Error: Output module: Trying to add a module to safety routing table which does not support FSoE.");
          LogHWPath("HW-Path of Module: {0}", pListHeader^.p_us_Path);
        end_if;
      else
        LogError("@0235 (SafetyBaseFSoE::AddModuleToRoutingTabs) Config Read Error: Output module: No Object of HW-class found for module to be added to safety routing table.");
        LogHWPath("HW-Path of Module: {0}", pListHeader^.p_us_Path);
      end_if;

    //add other cpu module

    elsif pModule = pListHeader then

      //the output module is addressed by the ListHeaderPath
      //get this-pointer of object in network that is located with transfered path
      MyPara.uiCmd := _BUS_IF_GET_OBJECT_THIS_PTR;
      MyPara.aPara[0] := pModule^.p_us_Path$DINT;
      sd_retval$iprStates := ToBusInterface.NewInst(#MyPara, #MyResult);
      p_TargetObject := MyResult.aData[0]$pVirtualBase;

      //this-pointer found
      if ( p_TargetObject ) then

        //check if it's a safety module
        MyPara.uiCmd := CMD_SM_GET_MODULE_TYPE;
        sd_retval$iprStates := p_TargetObject^.NewInst(#MyPara, #MyResult);

        if ( MyResult.aData[0]$UDINT = SM_TYPE_SAFETY_MODULE_FSOE ) then

          //object is based on SafetyBaseFSoE
          p_SafetyBase := p_TargetObject;

          //get safety number
          MyPara.uiCmd := CMD_SM_CONFIG_SAFETY_CPU;

          sd_retval$iprStates := p_SafetyBase^.NewInst(#MyPara, #MyResult);

          ud_IO_SafeNumber := MyResult.aData[0]$UDINT;

//          ud_IO_SafeNumber := p_SafetyBase^.ConfigSafetyCpu();

          if ( ud_IO_SafeNumber <> 0 ) then

            //add module to routing table
            sd_retval := AddRoutingElement( ud_SafeNumber       := ud_IO_SafeNumber
                                          , ud_thisp            := p_SafetyBase$UDINT
                                          , pObject             := pListHeader
                                          );
          elsif b_IsOptional = FALSE then
            LogError("@0236 (SafetyBaseFSoE::AddModuleToRoutingTabs) Config Read Error: CPU module: 0 is an invalid safety number.");
            LogHWPath("HW-Path of Module: {0}", pListHeader^.p_us_Path);

            b_ReInitMarker := TRUE;

          end_if;
        else
          LogError("@027E (SafetyBaseFSoE::AddModuleToRoutingTabs) Config Read Error: CPU module: Trying to add a module to safety routing table which does not support FSoE.");
          LogHWPath("HW-Path of Module: {0}", pListHeader^.p_us_Path);
        end_if;
      else
        LogError("@0238 (SafetyBaseFSoE::AddModuleToRoutingTabs) Config Read Error: CPU module: No Object of HW-class found for module to be added to safety routing table.");
        LogHWPath("HW-Path of Module: {0}", pListHeader^.p_us_Path);
      end_if;

    //add input module

    else
      //It's a safety input module, so it has to be added to safety input list.
      //check if found object represents a safety module
      MyPara.uiCmd := CMD_SM_GET_MODULE_TYPE;
      sd_retval$iprStates := p_TargetObject^.NewInst(#MyPara, #MyResult);
      if ( MyResult.aData[0]$UDINT = SM_TYPE_SAFETY_MODULE_FSOE ) then

        //object is based on SafetyBaseFSoE
        p_SafetyBase := p_TargetObject;

        //get safety number
        MyPara.uiCmd := CMD_SM_CONFIG_SAFETY_CPU;

        sd_retval$iprStates := p_SafetyBase^.NewInst(#MyPara, #MyResult);

        ud_IO_SafeNumber := MyResult.aData[0]$UDINT;

        //configure safety input module and receive pointer on PDO-Buffer and safety number
//        MyPara.uiCmd := CMD_SM_CONFIG_SAFETY_INPUT;
//        MyPara.aPara[0] := SafetyNumber$DINT;
//        MyPara.aPara[1] := this$DINT;
//        MyPara.aPara[2] := (#ud_PDO_Buffer)$DINT;
//        sd_retval$iprStates := p_SafetyBase^.NewInst(#MyPara, #MyResult);
//
//        ud_IO_SafeNumber := MyResult.aData[0]$UDINT;

//      ud_IO_SafeNumber := p_SafetyBase^.ConfigSafetyInput ( ud_SafeNrCPU    := SafetyNumber
//                                                          , ud_thisp        := this$UDINT
//                                                          , p_PDOBuffer     := #ud_PDO_Buffer
//                                                          , pMoveActive     := pMoveCommandInputActive
//                                                          , p_ud_MoveSourceAddr := #ud_MoveSourceAddr
//                                                          );

        //input module successfully configured
        if ( ud_IO_SafeNumber <> 0 ) then
(*
          // only if the configuration affects our cpu, we add something to our PDO input buffer
          MyPara.uiCmd := _BUS_IF_GET_OBJECT_THIS_PTR;
          MyPara.aPara[0] := pListHeader^.p_us_Path$DINT;
          sd_retval$iprStates := ToBusInterface.NewInst(#MyPara, #MyResult);
          p_TargetObject := MyResult.aData[0]$pVirtualBase;

//          p_TargetObject := ( GetObjectThisp(p_us_ObjectPath := pListHeader^.p_us_Path) )$pVirtualBase;

          //this-pointer found
          if ( p_TargetObject = this ) then

            //add pointer on PDO output buffer of input module to list of incoming PDOs
            sd_retval := AddPDOToInputBuffer(ud_p2Buffer         := ud_PDO_Buffer
                                           , ud_SafetyNr         := ud_IO_SafeNumber
                                           , b_IsOptional        := b_IsOptional
                                           );
          else
            sd_retval := 0;
          end_if;
*)
          if ( sd_retval = 0 ) then

            //add module to routing table
            sd_retval := AddRoutingElement( ud_SafeNumber       := ud_IO_SafeNumber
                                          , ud_thisp            := p_SafetyBase$UDINT
                                          , pObject             := pModule
                                          );

          else
            LogError("@0239 (SafetyBaseFSoE::AddModuleToRoutingTabs) Config Read Error: Input module: Failed to add module to input buffer.");
            LogHWPath("HW-Path of Module: {0}", pListHeader^.p_us_Path);
          end_if;
        else
          // module in configuration, which is not physically available but hw-class is placed
          sd_retval := 0; // could be an optional module
        end_if;
      else
        LogError("@027E (SafetyBaseFSoE::AddModuleToRoutingTabs) Config Read Error: Input module: Trying to add a module to safety routing table which does not support FSoE.");
        LogHWPath("HW-Path of Module: {0}", pModule^.p_us_Path);
      end_if;
    end_if;
  else
    // module in configuration, which is not physically available and no hw-class is placed
    LogError("@023B (SafetyBaseFSoE::AddModuleToRoutingTabs) Config Read Error: Module in safety configuration, where no HW-Class is placed (maybe optional module).");
    LogHWPath("HW-Path of Module: {0}", pModule^.p_us_Path);
    sd_retval := 0;
  end_if;

END_FUNCTION

FUNCTION VIRTUAL SafetyBaseFSoE::GetRoutingElementByThis
  VAR_INPUT
    ud_thisp 	: UDINT;
  END_VAR
  VAR_OUTPUT
    p_RoutElement 	: ^SafetyBaseFSoE::RoutElement;
  END_VAR
  VAR
    i1                  : UINT;
    p_RoutElement_Act   : ^RoutElement;
  END_VAR

  p_RoutElement := NIL;

  //set pointer on first routing element
  p_RoutElement_Act := p_RoutTable;

  //check each element
  for i1 := 0 to ui_CntRoutElements - 1 do

    //if searched this is found, pointer on routing element is returned
    if ( p_RoutElement_Act^.ud_Thisp = ud_thisp ) then
      p_RoutElement := p_RoutElement_Act;
      return;
    end_if;

    //set pointer to next element
    p_RoutElement_Act += sizeof ( RoutElement );

  end_for;

END_FUNCTION

FUNCTION VIRTUAL SafetyBaseFSoE::SDOStdRequ
  VAR_INPUT
    us_Command 	: USINT;
    p_us_RespData 	: ^USINT;
    us_RespLength 	: USINT;
  END_VAR
  VAR_OUTPUT
    sd_retval 	: DINT;
  END_VAR
  VAR
    pSDORequestBuffer   : ^t_SDOStdHeader;
    pSDOResponseBuffer  : ^SDOStdResp;
    RespBuffer          : ARRAY [0..127] OF USINT;
    RequBuffer          : ARRAY [0..127] OF USINT;
    us_OutLength        : USINT;
  END_VAR

  //SDO requests for this commands don't have any further data
  pSDORequestBuffer$^void := #RequBuffer[0];
  pSDOResponseBuffer$^void := #RespBuffer[0];

  //SDO response buffer (length header + rc + data)
  us_OutLength := sizeof(t_SDOStdHeader) + 1 + us_RespLength;

  //calculate length without crc
  pSDORequestBuffer^.len := sizeof(t_SDOStdHeader) - sizeof(t_SDOStdHeader.CRC);

  //type
  pSDORequestBuffer^.typ := SDO_STD;

  //sequence number
  pSDORequestBuffer^.SeqNr := us_CntSequNr;

  //increase counter for sequence number
  if us_CntSequNr < 16#7F then
    us_CntSequNr += 1;
  else
    us_CntSequNr := 0;
  end_if;

  //command to inform CPU about initializing classes is ok
  pSDORequestBuffer^.cmd := us_Command;

  //set CRC-field to 0
  pSDORequestBuffer^.CRC := 0;

  //send request
  sd_retval := SAFETY_iSendRequest( uiMaster    := 0
                                  , pucNode     := p_ObjectPath
                                  , uiInLength  := sizeof(t_SDOStdHeader)
                                  , pucInput    := pSDORequestBuffer$^USINT
                                  , uiOutLength := us_OutLength
                                  , pucOutput   := pSDOResponseBuffer$^USINT
                                  );

  //no response
  if ( sd_retval = 0 ) then

    //check sequence number to exclude a possible wrong response
    if ( pSDORequestBuffer^.SeqNr <> pSDOResponseBuffer^.StdHeader.SeqNr ) then
      sd_retval := -102;
      //log not routable SDOs
      LogValue("@022A (SafetyBaseFSoE::SDOStdRequ) Invalid Sequence number in SDO Standard Response. Got 0x{0} instead of expected 0x{1}", to_udint(pSDOResponseBuffer^.StdHeader.SeqNr), to_udint(pSDORequestBuffer^.SeqNr));

    //check returncode of SDO
    elsif ( pSDOResponseBuffer^.us_Returncode <> SBF_SDO_RETCODE_OK ) then
      //log not routable SDOs
      LogValue("@022B (SafetyBaseFSoE::SDOStdRequ) Safety module 0x{0}: Retcode of SDO Standard Response was invalid. Retcode: 0x{1}", SafetyNumber$UDINT, to_udint(pSDOResponseBuffer^.us_Returncode));
      sd_retval := -103;
    end_if;
  else
    //log not routable SDOs
    LogValue("@023E (SafetyBaseFSoE::SDOStdRequ) SAFETY_iSendRequest failed with retcode: -0x{0}", to_udint(ABS(sd_retval)));
  end_if;

  //return response
  if ( ( sd_retval = 0 ) & ( p_us_RespData <> NIL )) then

    ToStdLib.MemCpy(dest := p_us_RespData, source := #pSDOResponseBuffer^.us_Data, size := us_RespLength);

  end_if;

END_FUNCTION

FUNCTION VIRTUAL SafetyBaseFSoE::GetPDOInputBuffer
  VAR_INPUT
    ud_p2Buffer 	: UDINT;
    ud_SafetyNr 	: HDINT;
    p_FoundSafetyNr 	: ^BOOL;(* := NIL *)
    b_IsInterfaceFrame 	: BOOL;
    ui_TargetOffset 	: UINT;
  END_VAR
  VAR_OUTPUT
    p_InputBuffer 	: ^SafetyBaseFSoE::PDOInputBuffer;
  END_VAR
  VAR
    i1                : UINT;
    p_InputBuffer_Act : ^PDOInputBuffer;
  END_VAR

  p_InputBuffer := NIL;

  if p_FoundSafetyNr then
    p_FoundSafetyNr^ := FALSE;
  end_if;

  if ui_cnt_PDOInputBuffer then

    //set pointer on first input buffer element
    p_InputBuffer_Act := #aPDOInputBuffer[0];

    //check each element
    for i1 := 0 to (ui_cnt_PDOInputBuffer-1) do

      //if searched pointer is found, pointer on input buffer element is returned
      if (p_InputBuffer_Act^.ud_p2Buffer        = ud_p2Buffer )       &
         (p_InputBuffer_Act^.b_IsInterfaceFrame = b_IsInterfaceFrame) &

         // if it's an interface frame, the offset has to be the same (otherwise it could be a dynamically connected FlexCon)
        ((b_IsInterfaceFrame = FALSE) |
         (p_InputBuffer_Act^.ui_TargetOffset    = ui_TargetOffset))   then
        // even if found by SafetyNumber, if found by buffer => reset the found by safetynumber
        p_FoundSafetyNr^ := FALSE;
        p_InputBuffer := p_InputBuffer_Act;
        return;
      end_if;

      if p_FoundSafetyNr & (p_InputBuffer_Act^.ud_SafetyNr        = ud_SafetyNr)        &
                           (p_InputBuffer_Act^.b_IsInterfaceFrame = b_IsInterfaceFrame) &

                           // if it's an interface frame, the offset has to be the same (otherwise it could be a dynamically connected FlexCon)
                          ((b_IsInterfaceFrame = FALSE) |
                           (p_InputBuffer_Act^.ui_TargetOffset    = ui_TargetOffset))   then
        p_FoundSafetyNr^ := TRUE;
        p_InputBuffer := p_InputBuffer_Act;
//        return;
      end_if;

      //set pointer to next element
      p_InputBuffer_Act += sizeof ( PDOInputBuffer );

    end_for;
  end_if;

END_FUNCTION

FUNCTION VIRTUAL SafetyBaseFSoE::GetThisViaServerName
  VAR_INPUT
    pObjectDotServer 	: ^CHAR;
  END_VAR
  VAR_OUTPUT
    ThisPtr 	: ^void;
  END_VAR
  VAR
    ChannelMode : CHMODE;
  END_VAR

  ThisPtr := NIL;

  if pObjectDotServer = NIL then
    return;
  end_if;

  // get thispointer to server via name
  ChannelMode := _LookUpEmbed_C(pObjectDotServer, #ThisPtr, NIL);

  // check if it's a server
  case ChannelMode of
    _CH_CMD,
    _CH_SVR:

  else
    ThisPtr := NIL;
    LogError("@023F (SafetyBaseFSoE::GetThisViaServerName) Couldn't get thispointer of server:.");
    LogError(e_msg:=pObjectDotServer);
    ud_UnsafeVarsNotFound += 1;
  end_case;

END_FUNCTION

#pragma warning(disable: 73);
FUNCTION VIRTUAL SafetyBaseFSoE::LogError
  VAR_INPUT
    e_msg 	: ^CHAR;
  END_VAR

#ifdef HWC_LogError
  HWC_LogError(this, e_msg);
#endif

END_FUNCTION

FUNCTION VIRTUAL SafetyBaseFSoE::LogValue
  VAR_INPUT
    pString 	: ^CHAR;
    Value 	: UDINT;
    Value2 	: UDINT;(* := 16#FFFFFFFF *)
    Value3 	: UDINT;(* := 16#FFFFFFFF *)
  END_VAR

#ifdef HWC_LogValue3
  HWC_LogValue3(this, pString, Value, Value2, Value3);
#endif

END_FUNCTION
#pragma warning(default: 73);

FUNCTION VIRTUAL SafetyBaseFSoE::AddUnsafeRoutElement
  VAR_INPUT
    pRoutTable 	: ^SafetyBaseFSoE::pUnsafeIORoutingElement;
    pRoutElementsNo 	: ^UINT;
    ud_Address 	: UDINT;
    ui_NameLen 	: UINT;
    pNameNewElement 	: ^CHAR;
    BitMask 	: BDINT;(* := 0 *)
  END_VAR
  VAR_OUTPUT
    sd_retval 	: DINT;
  END_VAR
  VAR
    p_RoutElement   : ^UnsafeIORoutingElement;
    RemoteDomain      : USINT;
    LinearMemory : BOOL;
  END_VAR

  sd_retval := -1;

  // check parameters
  if (ui_NameLen = 0) | (pNameNewElement = NIL) then
    LogError("@0240 (SafetyBaseFSoE::AddUnsafeRoutElement) Invalid call parameters for the variable name (invalid configuration in safety cpu).");
    return;
  end_if;

  // on CSCP011 the SDO_COMMAND_WRITE_VALUES didn't exist, so we have to make a difference here
  if (pRoutTable = #p_UnsafeOutputsTable) then
    LinearMemory := TRUE;
  else
    LinearMemory := FALSE;
  end_if;

  // if there is a domain info attached
  if (pNameNewElement^ = '@') & ((pNameNewElement + 1)^ = 'D') then
    // check if it's in the actual domain
    if (pNameNewElement + 3)^ = ':' then
      // 1 digit domain number
      RemoteDomain := (pNameNewElement + 2)^ - '0';
    elsif (pNameNewElement + 4)^ = ':' then
      // 2 digits domain number
      RemoteDomain := ((pNameNewElement + 2)^ - '0') * 10 + (pNameNewElement + 3)^ - '0';
    else
      LogError("@0241 (SafetyBaseFSoE::AddUnsafeRoutElement) Invalid domain info at unsafe variable.");
      return;
    end_if;

    // prepare the string (remove the domain info)
    if RemoteDomain >= 10 then
      ui_NameLen -= 5;
      pNameNewElement += 5;
    else
      ui_NameLen -= 4;
      pNameNewElement += 4;
    end_if;
  end_if;

  //With the first element, the table must be positioned
  if ( pRoutTable^ = NIL ) then

    //allocate memory for first routing element
    pRoutTable^$^void := ToStdLib.Malloc(size := sizeof(UnsafeIORoutingElement));

    if ( pRoutTable^ = NIL ) then

      sd_retval                         := -1;
      SetSafetyState(NewState:=_MemAllocFailed);
      return;

    end_if;

    p_RoutElement := pRoutTable^;

  else

    //add new element

    //add space for one element to table (linked list element for inputs and linear data area for outputs)
    if LinearMemory = FALSE then
    // search for a place
      p_RoutElement := pRoutTable^;
      while p_RoutElement^.pNext do
        p_RoutElement := p_RoutElement^.pNext;
      end_while;
      p_RoutElement^.pNext$^void := ToStdLib.Malloc(sizeof(UnsafeIORoutingElement));

      if ( p_RoutElement^.pNext = NIL ) then

        sd_retval                         := -1;
        SetSafetyState(NewState:=_MemAllocFailed);
        return;

      end_if;

      // set pointer to new element
      p_RoutElement := p_RoutElement^.pNext;
    else
      pRoutTable^$^void := ToStdLib.ReAlloc(mptr := pRoutTable^, newsize := ( ( pRoutElementsNo^ + 1 ) * sizeof(UnsafeIORoutingElement)));

      if ( pRoutTable^ = NIL ) then

        sd_retval                         := -1;
        SetSafetyState(NewState:=_MemAllocFailed);
        return;

      end_if;

      //set pointer to empty element on last position
      p_RoutElement := pRoutTable^ + ( pRoutElementsNo^ ) * sizeof(UnsafeIORoutingElement);
    end_if;
  end_if;

  if p_RoutElement then
    //allocate memory for name
    p_RoutElement^.pName$^void := ToStdLib.Malloc(size := ui_NameLen);

    if ( p_RoutElement^.pName = NIL ) then

      sd_retval                         := -1;
      SetSafetyState(NewState:=_MemAllocFailed);
      return;

    end_if;

    p_RoutElement^.NameLength := ui_NameLen;
    _memcpy(ptr1:=p_RoutElement^.pName, ptr2:=pNameNewElement, cntr:=ui_NameLen);

    // unsafe bdint variables are localized in a different memory area
    if BitMask then
      p_RoutElement^.ud_Address := SBF_SDO_ADDRESS_UNSAFE_BDINT + ud_Address;
    else
      p_RoutElement^.ud_Address := SBF_SDO_ADDRESS_APP_DATA + ud_Address;
    end_if;

    p_RoutElement^.BitMask := BitMask;

    // initialize with invalid
    p_RoutElement^.b_IsValid            := FALSE;
    p_RoutElement^.sd_OldValue          := (16#80000000)$DINT;
    p_RoutElement^.sd_NewValue4External := (16#80000000)$DINT;

    // remember that we haven't transmitted this value so far
    p_RoutElement^.b_AlreadyTransmitted := FALSE;

    // initialize next pointer
    p_RoutElement^.pNext := NIL;

    //increase counter
    pRoutElementsNo^ += 1;

    // check if name exists in PLC
    p_RoutElement^.ud_Thisp   := GetThisViaServerName(pNameNewElement)$UDINT;
    if (pRoutTable = #p_UnsafeOutputsTable) & p_RoutElement^.BitMask then
      p_RoutElement^.UnsafeType := BDINTOutput;
    else
      p_RoutElement^.UnsafeType := NormalUnsafe;
    end_if;
  end_if;

END_FUNCTION

FUNCTION VIRTUAL SafetyBaseFSoE::InitPathInfo
  VAR_INPUT
    pPathInfo 	: ^SafetyBaseFSoE::PathInfoType;
  END_VAR

  pPathInfo^.p_us_Path := NIL;
  pPathInfo^.p_us_PathComp := NIL;
  pPathInfo^.ui_PathCompLen := 0;

END_FUNCTION

FUNCTION VIRTUAL SafetyBaseFSoE::ResetConfig
  VAR
    p_SafetyBase        : pVirtualBase;
    p_RoutElement       : ^RoutElement;
    p_UnsafeRoutElement : ^UnsafeIORoutingElement;
    i                   : UINT;
    MyPara              : CmdStruct;
    MyResult            : results;
  END_VAR

  // tell all modules, which are connected to this cpu (through the old configuration) that they should delete the cpu from their routing table
  // must be more than 1, because 1st is always own entry
  if p_RoutTable & (ui_CntRoutElements > 1) then
    //set pointer on 2nd routing element
    p_RoutElement := p_RoutTable + sizeof(RoutElement);
    for i := 1 to (ui_CntRoutElements - 1) do
      // clear everything except this object (done after the for loop)
      if p_RoutElement^.ud_Thisp <> THIS$UDINT then
        // get thispointer of routing element
        p_SafetyBase := (p_RoutElement^.ud_Thisp)$pVirtualBase;

        // call other safety-class to remove the safetynumber from the routing table
        MyPara.uiCmd := CMD_SM_REMOVE_CPU_FROM_TABLE;
        MyPara.aPara[0] := SafetyNumber$DINT;

        p_SafetyBase^.NewInst(#MyPara, #MyResult);

//        p_SafetyBase^.RemoveCPUFromTable(ud_SafetyNr := SafetyNumber);
      end_if;

      // free memory of compressed path
      if p_RoutElement^.p_CompressedPath then
        ToStdLib.Free(mptr:=p_RoutElement^.p_CompressedPath);
      end_if;

      // set pointer on next routing element
      p_RoutElement += sizeof(RoutElement);
    end_for;

    // reduce local routing table to the cpu's own entry
    ui_CntRoutElements := 1;
  end_if;

  // on CSCP011 the SDO_COMMAND_WRITE_VALUES didn't exist, so we have to make a difference here
  while p_UnsafeInputsTable do
    p_UnsafeRoutElement := p_UnsafeInputsTable;
    p_UnsafeInputsTable := p_UnsafeInputsTable^.pNext;

    ToStdLib.Free(mptr:=p_UnsafeRoutElement^.pName);
    ToStdLib.Free(mptr:=p_UnsafeRoutElement);
  end_while;
  ui_CntUnsafeInputs := 0;

  // unsafe outputs are always in linear memory
  if p_UnsafeOutputsTable then
    ToStdLib.Free(mptr:=p_UnsafeOutputsTable);
    p_UnsafeOutputsTable := NIL;
  end_if;
  ui_CntUnsafeOutputs := 0;

  // reset no of SDO input buffer
  ui_cnt_SDOInputBuffer := 0;

  // if the old configuration is reset, check for the configured state of the cpu
  b_CheckConfigured := TRUE;

END_FUNCTION

FUNCTION VIRTUAL SafetyBaseFSoE::RemoveCPUFromTable
  VAR_INPUT
    ud_SafetyNr 	: HDINT;
  END_VAR
  VAR
    p_RoutElement   : ^RoutElement;
    i               : UDINT;
    FoundIndex      : UDINT;
    pPDOInputBuffer : ^PDOInputBuffer;
    Found : BOOL;
  END_VAR

  // if we are a cpu, do nothing
  if b_CheckCRC then
    return;
  end_if;

  //check each element (must be more than 1, because 1st is always own entry)
  if p_RoutTable & (ui_CntRoutElements > 1) then
    //set pointer on 2nd routing element
    p_RoutElement := p_RoutTable + sizeof(RoutElement);
    for i := 1 to (ui_CntRoutElements - 1) do

      // if we found safenumber, delete element from table
      if ( p_RoutElement^.ud_SafeNumber = ud_SafetyNr ) then

        // at last element we don't need to copy data, just decrease buffersize
        if i <> (ui_CntRoutElements - 1) then
          _memcpy(p_RoutElement, p_RoutElement + sizeof(RoutElement), sizeof(RoutElement) * (ui_CntRoutElements - 1 - i));
        end_if;

        // free 1 element and decrease element counter
        ui_CntRoutElements -= 1;

        exit;
      end_if;

      // set pointer on next routing element
      p_RoutElement += sizeof(RoutElement);
    end_for;
  end_if;

  // reset no of SDO input buffer
  ui_cnt_SDOInputBuffer := 0;

  // check if we received a PDO from this CPU => if so, delete it from the PDO input buffer
  if ui_cnt_PDOInputBuffer then
    // search for the PDO
    Found := FALSE;
    pPDOInputBuffer := #aPDOInputBuffer[0];
    for FoundIndex := 0 to (ui_cnt_PDOInputBuffer-1) do
      if pPDOInputBuffer^.ud_SafetyNr = ud_SafetyNr then
        Found := TRUE;
        exit;
      end_if;

      pPDOInputBuffer += sizeof(PDOInputBuffer);
    end_for;

    // if we found the PDO => remove it from memory (move the memory behind the found PDO over the place of the found PDO)
    if Found then
      // if it's last entry (no entries have to be moved) => we only have to copy some memory if it's not the last
      if FoundIndex < (ui_cnt_PDOInputBuffer-1) then
        for i := FoundIndex to (ui_cnt_PDOInputBuffer-2) do
          aPDOInputBuffer[i] := aPDOInputBuffer[i+1];
        end_for;
      end_if;
      ui_cnt_PDOInputBuffer -= 1;

      if ui_cnt_PDOInputBuffer = 0 then
        if ModuleSyncNo & (SafetyState <> _SafetyClassOK) then
          ModuleSyncNo -= 1;
        end_if;
      end_if;
    end_if;
  end_if;

END_FUNCTION

FUNCTION VIRTUAL SafetyBaseFSoE::CheckUnsafeUpdateCycle

  // we can only use 56 byte pay load (instead of 64) because fw drops the 8 byte used for addresses in safe SDO

  if ui_CntUnsafeOutputs then
  // maximum of read variables in 1 frame is 15 (56 Bytes pay load - 1 Byte Returncode - 1 Byte Length = 54 Bytes => 13x4Bytes = 52)
    MaxVarsPerReadPackage := (SBF_SDO_MAX_LENGTH - (sizeof(SDOHeader) - sizeof(SDOHeader.SessId)) - sizeof(SDORespReadConfig.us_Returncode) - sizeof(SDORespReadConfig.us_Length)) / sizeof(DINT);
    ReadFramesNeeded := ((ui_CntUnsafeOutputs - 1) / MaxVarsPerReadPackage) + 1;
  else
    ReadFramesNeeded := 0;
  end_if;

  if ui_CntUnsafeInputs then
  // maximum of write variables in 1 frame is 14 (56 Bytes pay load - 4 Byte Address - 1 Byte Length = 51 Bytes => 12x4Bytes = 48)
    MaxVarsPerWritePackage := (SBF_SDO_MAX_LENGTH - (sizeof(SDOHeader) - sizeof(SDOHeader.SessId)) - sizeof(SDORequReadConfig.ud_Address) - sizeof(SDORequReadConfig.us_Length)) / sizeof(DINT);
    WriteFramesNeeded := ((ui_CntUnsafeInputs - 1) / MaxVarsPerWritePackage) + 1;
  else
    WriteFramesNeeded := 0;
  end_if;

  // check if user has given us enough time
  ud_TransfertimePerPackage := SBF_SDO_TRANSFERTIME;

  if ( (WriteFramesNeeded + ReadFramesNeeded) * ud_TransfertimePerPackage ) > ServerUpdateTime then
    ServerUpdateTime := ( WriteFramesNeeded + ReadFramesNeeded ) * ud_TransfertimePerPackage;
    ud_ServerUpdateTime := ( ReadFramesNeeded ) * ud_TransfertimePerPackage;
  end_if;

END_FUNCTION

FUNCTION VIRTUAL GLOBAL SafetyBaseFSoE::FetchDiagState

  DiagVars.UserDiagStateReady := FALSE;
  DiagVars.UserWantsDiagState := TRUE;

END_FUNCTION

FUNCTION VIRTUAL GLOBAL SafetyBaseFSoE::GetDiagState
  VAR_INPUT
    pDiagState 	: ^SafetyDiagState;
  END_VAR
  VAR_OUTPUT
    StateReady 	: BOOL;
  END_VAR

  StateReady := DiagVars.UserDiagStateReady;

  // if data ready, we save it into user structure
  if StateReady then
    pDiagState^.RunState            := DiagVars.UserGetStateResp.RuntimeState;
    pDiagState^.ConfigState         := DiagVars.UserGetStateResp.ConfigState;
    pDiagState^.LoginLevel          := DiagVars.UserGetStateResp.LoginLevel;
    pDiagState^.ErrorCounterIOState := DiagVars.UserGetStateResp.ErrorCount;
  end_if;

END_FUNCTION

FUNCTION VIRTUAL GLOBAL SafetyBaseFSoE::FetchDiagInfo
  VAR_INPUT
    ucChoice 	: USINT;
  END_VAR

  DiagVars.ucChoiceDiagInfo  := ucChoice;
  DiagVars.UserDiagInfoReady := FALSE;
  DiagVars.UserWantsDiagInfo := TRUE;

END_FUNCTION

FUNCTION VIRTUAL GLOBAL SafetyBaseFSoE::GetDiagInfo
  VAR_INPUT
    pDiagInfo 	: ^SafetyDiagInfo;
  END_VAR
  VAR_OUTPUT
    StateReady 	: BOOL;
  END_VAR

  StateReady := DiagVars.UserDiagInfoReady;

  // if data ready, we save it into user structure
  if StateReady then
    pDiagInfo^ := DiagVars.UserGetDiagInfoResp;
  end_if;

END_FUNCTION

FUNCTION VIRTUAL SafetyBaseFSoE::SDORequ
  VAR_INPUT
    us_Command 	: USINT;
    p_us_RequData 	: ^USINT;
    us_RequLength 	: USINT;
    p_us_RespData 	: ^USINT;
    us_RespLength 	: USINT;
  END_VAR
  VAR_OUTPUT
    sd_retval 	: DINT;
  END_VAR
  VAR
    pSDORequestBuffer   : ^t_SDOStdHeader;
    pSDOResponseBuffer  : ^SDOStdResp;
    RespBuffer          : ARRAY [0..127] OF USINT;
    RequBuffer          : ARRAY [0..127] OF USINT;
    us_InLength         : USINT;
    us_OutLength        : USINT;
  END_VAR

  //SDO requests for this commands don't have any further data
  pSDORequestBuffer$^void := #RequBuffer[0];
  pSDOResponseBuffer$^void := #RespBuffer[0];

  //SDO request buffer (length header + data)
  us_InLength := sizeof(t_SDOStdHeader) + us_RequLength;

  //SDO response buffer (length header + rc + data)
  us_OutLength := sizeof(t_SDOStdHeader) + 1 + us_RespLength;

  //calculate length without crc
  pSDORequestBuffer^.len := sizeof(t_SDOStdHeader) - sizeof(t_SDOStdHeader.CRC) + us_RequLength;

  //type
  pSDORequestBuffer^.typ := SDO_STD;

  //sequence number
  pSDORequestBuffer^.SeqNr := us_CntSequNr;

  _memcpy(ptr1:=pSDORequestBuffer + sizeof(t_SDOStdHeader), ptr2:=p_us_RequData, cntr:=us_RequLength);

  //increase counter for sequence number
  if us_CntSequNr < 16#7F then
    us_CntSequNr += 1;
  else
    us_CntSequNr := 0;
  end_if;

  //command to inform CPU about initializing classes is ok
  pSDORequestBuffer^.cmd := us_Command;

  //set CRC-field to 0
  pSDORequestBuffer^.CRC := 0;

  //send request
  sd_retval := SAFETY_iSendRequest( uiMaster    := 0
                                  , pucNode     := p_ObjectPath
                                  , uiInLength  := us_InLength
                                  , pucInput    := pSDORequestBuffer$^USINT
                                  , uiOutLength := us_OutLength
                                  , pucOutput   := pSDOResponseBuffer$^USINT
                                  );

  //no response
  if ( sd_retval = 0 ) then

    //check sequence number to exclude a possible wrong response
    if ( pSDORequestBuffer^.SeqNr <> pSDOResponseBuffer^.StdHeader.SeqNr ) then
      sd_retval := -102;

    //check returncode of SDO
    elsif ( pSDOResponseBuffer^.us_Returncode <> SBF_SDO_RETCODE_OK ) then
      sd_retval := -103;
    end_if;

  end_if;

  //return response
  if ( ( sd_retval = 0 ) & ( p_us_RespData <> NIL )) then
    ToStdLib.MemCpy(dest := p_us_RespData, source := #pSDOResponseBuffer^.us_Data, size := us_RespLength);
  end_if;

END_FUNCTION

FUNCTION VIRTUAL GLOBAL SafetyBaseFSoE::SaveLog
  VAR_INPUT
    ucChoice 	: USINT;
    pDPNE 	: ^CHAR;
  END_VAR
  VAR_OUTPUT
    Success 	: DINT;
  END_VAR

  if DiagVars.SavingLogInProgress = FALSE then
    DiagVars.SavingLogInProgress := TRUE;

    DiagVars.SavingLogSuccessful := FALSE; //Reset Value

    DiagVars.ucChoiceSaveLog := ucChoice;

    _memcpy(ptr1:=#DiagVars.DPNE, ptr2:=pDPNE, cntr:=_strlen(pDPNE));

    Success := TRUE;
  else
    Success := FALSE;
  end_if;

END_FUNCTION

FUNCTION VIRTUAL GLOBAL SafetyBaseFSoE::SaveLogActive
  VAR_OUTPUT
    InProgress 	: BOOL;
  END_VAR

  InProgress := DiagVars.SavingLogInProgress;

END_FUNCTION

FUNCTION VIRTUAL SafetyBaseFSoE::BlockedTransferLength
  VAR_INPUT
    ud_Datalength 	: UDINT;
    us_MaxBlocklength 	: USINT;
  END_VAR
  VAR_OUTPUT
    us_ActBlocklength 	: USINT;
  END_VAR

  IF ud_Datalength > to_UDINT(us_MaxBlocklength) THEN
    us_ActBlocklength := us_MaxBlocklength;
  ELSE
    us_ActBlocklength := to_USINT(ud_Datalength);
  END_IF;

END_FUNCTION

#pragma warning(disable: 73)
FUNCTION VIRTUAL SafetyBaseFSoE::AddFrame
  VAR_INPUT
    pFrame 	: ^t_SDOStdHeader;
    FrameState 	: DINT;
    CallerSafetyNr 	: HDINT;
  END_VAR

END_FUNCTION
#pragma warning(default: 73)

FUNCTION VIRTUAL SafetyBaseFSoE::RecordFrame
  VAR_INPUT
    pFrame 	: ^DINT;
    FrameState 	: DINT;
    IsFSoEPDO 	: BOOL;(* := FALSE *)
  END_VAR
  VAR
    ThisBackup  : pVoid;
    TempSafetyNr: HDINT;
    Length      : USINT;
  END_VAR

  if pAnalyzerThis & pAnalyzerMethod then

    TempSafetyNr := SafetyNumber;

    if IsFSoEPDO then

      // if write
      if FrameState then
        if aWritePDOs[0].Length > sizeof(PDOType.DataAndCopy) then
          Length := sizeof(PDOType.DataAndCopy);
        else
          Length := aWritePDOs[0].Length;
        end_if;

        // if it's the same content as last time
        if (_memcmp(ptr1:=pFrame, ptr2:=#OldFakePDOWrite.DataAndCopy[0], cntr:=Length) = 0) then
          // don't record it
          return;
        end_if;

        // fake the header
        OldFakePDOWrite.Length              := sizeof(PDOType) - sizeof(PDOType.CRC) - sizeof(PDOType.DataAndCopy) + Length;
        OldFakePDOWrite.FrameType.PDO       := TRUE;
        OldFakePDOWrite.FrameType.Reserved2 := TRUE;

        // store the PDO data (remember it as the last recorded)
        _memcpy(ptr1:=#OldFakePDOWrite.DataAndCopy[0], ptr2:=pFrame, cntr:=Length);

        pFrame := (#OldFakePDOWrite)$^DINT;

      // if read
      else
        if aReadPDOs[0].Length > sizeof(PDOType.DataAndCopy) then
          Length := sizeof(PDOType.DataAndCopy);
        else
          Length := aReadPDOs[0].Length;
        end_if;

        // if it's the same content as last time
        if (_memcmp(ptr1:=pFrame, ptr2:=#OldFakePDORead.DataAndCopy[0], cntr:=Length) = 0) then
          // don't record it
          return;
        end_if;

        // fake the header
        OldFakePDORead.Length              := sizeof(PDOType) - sizeof(PDOType.CRC) - sizeof(PDOType.DataAndCopy) + Length;
        OldFakePDORead.FrameType.PDO       := TRUE;
        OldFakePDORead.FrameType.Reserved2 := TRUE;

        // store the PDO data (remember it as the last recorded)
        _memcpy(ptr1:=#OldFakePDORead.DataAndCopy[0], ptr2:=pFrame, cntr:=Length);

        pFrame := (#OldFakePDORead)$^DINT;
      end_if;
    end_if;

    ThisBackup := THIS;

    THIS := pAnalyzerThis$^SafetyBaseFSoE;
    pAnalyzerMethod$AddFrame(pFrame$^t_SDOStdHeader, FrameState, TempSafetyNr);

    THIS := ThisBackup$^SafetyBaseFSoE;
  end_if;

END_FUNCTION

FUNCTION VIRTUAL SafetyBaseFSoE::ShowProjectRevision

// overload this for CPU modules

END_FUNCTION

FUNCTION SafetyBaseFSoE::DOCheck
  VAR_INPUT
    pFrame 	: ^t_SDOStdHeader;
    pCheckStruct 	: ^SafetyBaseFSoE::t_DataObjectCheck;
  END_VAR
  VAR
    DOCheckHeader : t_SDOStdHeader;
    ActTime : UDINT;
  END_VAR

  // check if input parameters are correct
  if pFrame & pFrame^.Len & pCheckStruct then
    DOCheckHeader := pFrame^;

    // only if we got a different frame
    if DOCheckHeader <> pCheckStruct^.LastHeader then
      ActTime := OS_READMICROSEC();

      pCheckStruct^.TimeDiff := ActTime - pCheckStruct^.LastTime;

      if pCheckStruct^.TimeDiff > pCheckStruct^.TimeDiffMax then
        if pCheckStruct^.TimeDiffMax = 0 then
          pCheckStruct^.TimeDiffMax := 1;
        else
          pCheckStruct^.TimeDiffMax := pCheckStruct^.TimeDiff;
        end_if;
      end_if;

      if pCheckStruct^.TimeDiff < pCheckStruct^.TimeDiffMin then
        pCheckStruct^.TimeDiffMin := pCheckStruct^.TimeDiff;
      end_if;

      pCheckStruct^.LastTime := ActTime;
    else
      // if it's the same frame again: problem!
      pCheckStruct^.SameFrameCnt += 1;
    end_if;
    pCheckStruct^.LastHeader := DOCheckHeader;
  end_if;

END_FUNCTION

FUNCTION VIRTUAL SafetyBaseFSoE::CalcPDOLength
  VAR_INPUT
    BoolVarNo 	: UDINT;
    DintVarNo 	: UDINT;
  END_VAR
  VAR_OUTPUT
    PdoLen 	: USINT;
  END_VAR
  VAR
    PayLoad : USINT;
  END_VAR

  // we have at least the header
  PdoLen := sizeof(PDOType) - sizeof(PDOType.DataAndCopy);
  PayLoad := 0;

  // now add some space for the needed data
  if BoolVarNo then
    // 1 byte (type + number of values) + 1 byte index + 2 bits for every value (4 per byte)
    PayLoad += 2 + ((BoolVarNo$USINT + 3) / 4);

    // make the it 2 byte aligned (if it isn't already) => only if no dint variables, otherwise it is done one at the DINT variables
    if (PayLoad MOD 2) & (DintVarNo = 0) then
      PayLoad := PayLoad + (2 - (PayLoad MOD 2)); //increase memory, up to a value, which could be divided by 2
    end_if;
  end_if;

  if DintVarNo then
    // 1 byte (type + number of values) + 1 byte index + 1 byte errorflags per 8 values + 4 byte for every value
    PayLoad += 2 + (((DintVarNo$USINT - 1 ) / 8) + 1) + DintVarNo$USINT * 4;

    // make the it 2 byte aligned (if it isn't already)
    if (PayLoad MOD 2) then
      PayLoad := PayLoad + (2 - (PayLoad MOD 2)); //increase memory, up to a value, which could be divided by 2
    end_if;
  end_if;

  // duplicate it
  PayLoad *= 2;

  // add it to the total length
  PdoLen += PayLoad;

END_FUNCTION

FUNCTION VIRTUAL SafetyBaseFSoE::AddModuleToCfg
  VAR_INPUT
    ModuleCfg 	: t_ModuleCfg;
  END_VAR
  VAR_OUTPUT
    retcode 	: DINT;
  END_VAR
  VAR
    pHelp : ^t_ModuleListElem;
  END_VAR

  retcode := 0;

  if pFirstModuleCfg = NIL then
    pFirstModuleCfg$pVoid := ToStdLib.Malloc(size:=sizeof(t_ModuleListElem));
    pHelp := pFirstModuleCfg;
  else
    pHelp := pFirstModuleCfg;
    // if searched path has been found, we already got this module in our list
    if (ModuleCfg.PathLen = pHelp^.ModuleInfo.PathLen) & (ToStdLib.MemCmp(dest:= ModuleCfg.pPath, source:= pHelp^.ModuleInfo.pPath , size:= ModuleCfg.PathLen) = 0) then
      // already in buffer => leave function
      return;
    end_if;
    while pHelp^.pNext <> NIL do
      // if searched path has been found, we already got this module in our list
      if (ModuleCfg.PathLen = pHelp^.ModuleInfo.PathLen) & (ToStdLib.MemCmp(dest:= ModuleCfg.pPath, source:= pHelp^.ModuleInfo.pPath , size:= ModuleCfg.PathLen) = 0) then
        // already in buffer => leave function
        return;
      else
        pHelp := pHelp^.pNext;
      end_if;
    end_while;

    // if searched path has been found, we already got this module in our list
    if (ModuleCfg.PathLen = pHelp^.ModuleInfo.PathLen) & (ToStdLib.MemCmp(dest:= ModuleCfg.pPath, source:= pHelp^.ModuleInfo.pPath , size:= ModuleCfg.PathLen) = 0) then
      // already in buffer => leave function
      return;
    else
      pHelp^.pNext$pvoid := ToStdLib.Malloc(size:=sizeof(t_ModuleListElem));
      pHelp := pHelp^.pNext;
    end_if;
  end_if;

  if pHelp <> NIL then
    // allocate memory for the module path
    pHelp^.ModuleInfo.pPath$pVoid := ToStdLib.Malloc(size:=ModuleCfg.PathLen);
    if pHelp^.ModuleInfo.pPath = NIL then
      SetSafetyState(NewState:=_MemAllocFailed);
      retcode := -1;
      return;
    end_if;

    _memcpy(ptr1:=pHelp^.ModuleInfo.pPath, ptr2:=ModuleCfg.pPath, cntr:=ModuleCfg.PathLen);

    // allocate memory for the module path
    pHelp^.ModuleInfo.pCompPath$pVoid := ToStdLib.Malloc(size:=ModuleCfg.CompPathLen);
    if pHelp^.ModuleInfo.pCompPath = NIL then
      SetSafetyState(NewState:=_MemAllocFailed);

      retcode := -1;
      return;
    end_if;

    _memcpy(ptr1:=pHelp^.ModuleInfo.pCompPath, ptr2:=ModuleCfg.pCompPath, cntr:=ModuleCfg.CompPathLen);

    pHelp^.ModuleInfo.Info        := ModuleCfg.Info;
    pHelp^.ModuleInfo.SafetyNbr   := ModuleCfg.SafetyNbr;
    pHelp^.ModuleInfo.InterfaceCRC:= ModuleCfg.InterfaceCRC;
    pHelp^.ModuleInfo.DestCRCNo   := ModuleCfg.DestCRCNo;
    phelp^.ModuleInfo.pDestCRCs   := ModuleCfg.pDestCRCs;
    pHelp^.ModuleInfo.PathLen     := ModuleCfg.PathLen;
    pHelp^.ModuleInfo.CompPathLen := ModuleCfg.CompPathLen;
    pHelp^.ModuleInfo.PdoOutLen   := ModuleCfg.PdoOutLen;

    pHelp^.pNext                  := NIL;

    ModuleCfgNo += 1;
  else
    SetSafetyState(NewState:=_MemAllocFailed);
    retcode := -1;
    return;
  end_if;

END_FUNCTION

FUNCTION VIRTUAL SafetyBaseFSoE::AddPdoToCfg
  VAR_INPUT
    PdoCfg 	: t_PdoCfg;
  END_VAR
  VAR_OUTPUT
    retcode 	: DINT;
  END_VAR
  VAR
    pHelp : ^t_PdoListElem;
  END_VAR
//#pragma message("RamAnd 04.11.2014 17:18 \ die Aufrufe dieser Methode wurden unterbunden, da diese PDO-Infos für FSoE keine Relevanz haben")

  retcode := 0;

  if pFirstPdoCfg = NIL then
    pFirstPdoCfg$pVoid := ToStdLib.Malloc(size:=sizeof(t_PdoListElem));
    pHelp := pFirstPdoCfg;
  else
    pHelp := pFirstPdoCfg;
    // if searched path has been found, we already got this pdo in our list
    if (PdoCfg.SourcePathLen = pHelp^.PdoInfo.SourcePathLen) & (PdoCfg.DestPathLen = pHelp^.PdoInfo.DestPathLen) &
      (PdoCfg.InterfaceCRC = pHelp^.PdoInfo.InterfaceCRC) &
      (ToStdLib.MemCmp(dest:= PdoCfg.pSourcePath, source:= pHelp^.PdoInfo.pSourcePath , size:= PdoCfg.SourcePathLen) = 0) &
      (ToStdLib.MemCmp(dest:= PdoCfg.pDestPath,   source:= pHelp^.PdoInfo.pDestPath   , size:= PdoCfg.DestPathLen  ) = 0) then
      // already in buffer => leave function
      return;
    end_if;
    while pHelp^.pNext <> NIL do
      // if searched path has been found, we already got this pdo in our list
      if (PdoCfg.SourcePathLen = pHelp^.PdoInfo.SourcePathLen) & (PdoCfg.DestPathLen = pHelp^.PdoInfo.DestPathLen) &
        (PdoCfg.InterfaceCRC = pHelp^.PdoInfo.InterfaceCRC) &
        (ToStdLib.MemCmp(dest:= PdoCfg.pSourcePath, source:= pHelp^.PdoInfo.pSourcePath , size:= PdoCfg.SourcePathLen) = 0) &
        (ToStdLib.MemCmp(dest:= PdoCfg.pDestPath,   source:= pHelp^.PdoInfo.pDestPath   , size:= PdoCfg.DestPathLen  ) = 0) then
        // already in buffer => leave function
        return;
      else
        pHelp := pHelp^.pNext;
      end_if;
    end_while;
